// POUs/_FB_VisuDelta
(****************************************************************************************************<br>
© Syntegon Group.<br>
All rights reserved, also regarding any disposal, exploitation, reproduction, editing, distribution,<br>
as well as in the event of applications for industrial property rights.<br>
*****************************************************************************************************<br>
DESCRIPTION:<br>
One visualised Delta robot. Typical cycle:<br>
  fb_Delta.m_Register(vio_Manifest := GVL_Visu.stManifest, vi_udn_Id := 10, vi_str_Name := 'Delta 1',<br>
      vi_str_Path := 'MAIN.fb_Delta.vo_Visu');<br>
  fb_Delta.m_Configure(vi_Pose := BasePose, vi_lr_BaseRadius := 200, vi_lr_EffectorRadius := 50,<br>
      vi_lr_UpperArmLength := 400, vi_lr_LowerArmLength := 1000);<br>
  fb_Delta.m_SetFinger(vi_un_Finger := 1, vi_lr_Diameter := 40, vi_lr_Height := 50);<br>
  fb_Delta.m_SetWorkingArea(vi_lr_Radius := 750, vi_lr_ZMin := -1300, vi_lr_ZMax := -700, vi_lr_ConeHeight := 200,<br>
      vi_lr_ConeBottomRadius := 450);<br>
  fb_Delta.m_SetLimitArea(vi_lr_XMin := -500, vi_lr_XMax := 500, vi_lr_YMin := -750, vi_lr_YMax := 750,<br>
      vi_lr_ZMin := -1500, vi_lr_ZMax := -700);<br>
  fb_Delta.m_SetZone(vi_un_Zone := 1, vi_udn_ConveyorId := 1, vi_lr_Start := 1100, vi_lr_End := 1900,<br>
      vi_lr_AllocationOffset := 300);<br>
  fb_Delta.m_SetTcp(vi_ActualTcp := ActualTcp, vi_SetpointTcp := SetpointTcp);<br>
  fb_Delta.m_SetFingerState(vi_un_Finger := 1, vi_Pose := CupPose, vi_b_Active := b_Vacuum);<br>
Only the TCP (the gripper flange) is reported; the visualisation derives the arms from it. Tool rotations<br>
(e.g. a 4th axis) show only through the finger poses, absolute in the MCS. The config methods may be called<br>
every cycle; the config version only changes when a value does.<br>
*****************************************************************************************************<br>
OUTPUT VALUES:<br>
vo_Visu is the contract structure the gateway reads at the path given to m_Register. Do not write it.<br>
*****************************************************************************************************<br>
VERSION         ¦ DATE       ¦ NAME      ¦ CHANGE<br>
Syn_Visu 3.0.0  ¦ 2026-10-31 ¦ J.Willner ¦ Naming and layout after the TCAT programming guideline<br>
Syn_Visu 4.0.0  ¦ 2026-11-01 ¦ J.Willner ¦ Zones and fingers from _FB_VisuRobot; m_SetZone by index, no kind<br>
****************************************************************************************************)
FUNCTION_BLOCK _FB_VisuDelta EXTENDS _FB_VisuRobot
VAR_OUTPUT
	vo_Visu								: ST_VisuDelta;	// contract structure read by the gateway
END_VAR

(****************************************************************************************************<br>
© Syntegon Group.<br>
All rights reserved, also regarding any disposal, exploitation, reproduction, editing, distribution,<br>
as well as in the event of applications for industrial property rights.<br>
*****************************************************************************************************<br>
DESCRIPTION:<br>
Takes over vio_New and increments the config version if it differs from the current config. TRUE if changed.<br>
****************************************************************************************************)
METHOD PRIVATE m_ApplyConfig : BOOL
VAR_IN_OUT
	vio_New								: ST_VisuDeltaConfig;
END_VAR
m_ApplyConfig := Tc2_System.MEMCMP(ADR(vio_New), ADR(vo_Visu.stConfig), SIZEOF(vio_New)) <> 0;
IF m_ApplyConfig THEN
	vo_Visu.stConfig := vio_New;
	m_NotifyConfigChanged();
END_IF
END_METHOD

(****************************************************************************************************<br>
© Syntegon Group.<br>
All rights reserved, also regarding any disposal, exploitation, reproduction, editing, distribution,<br>
as well as in the event of applications for industrial property rights.<br>
*****************************************************************************************************<br>
DESCRIPTION:<br>
Base pose last set by m_Configure, MCS.<br>
****************************************************************************************************)
METHOD m_BasePose : ST_VisuPose
m_BasePose := vo_Visu.stConfig.stPose;
END_METHOD

(****************************************************************************************************<br>
© Syntegon Group.<br>
All rights reserved, also regarding any disposal, exploitation, reproduction, editing, distribution,<br>
as well as in the event of applications for industrial property rights.<br>
*****************************************************************************************************<br>
DESCRIPTION:<br>
Removes the limit area. TRUE if changed.<br>
****************************************************************************************************)
METHOD m_ClearLimitArea : BOOL
VAR
	TempNew								: ST_VisuDeltaConfig;
	TempEmpty							: ST_VisuLimitArea;
END_VAR
TempNew := vo_Visu.stConfig;
TempNew.stLimitArea := TempEmpty;
m_ClearLimitArea := m_ApplyConfig(TempNew);
END_METHOD

(****************************************************************************************************<br>
© Syntegon Group.<br>
All rights reserved, also regarding any disposal, exploitation, reproduction, editing, distribution,<br>
as well as in the event of applications for industrial property rights.<br>
*****************************************************************************************************<br>
DESCRIPTION:<br>
Manifest type: Delta robot.<br>
****************************************************************************************************)
METHOD PROTECTED m_ComponentType : E_VisuComponentType
m_ComponentType := E_VisuComponentType.DELTA;
END_METHOD

(****************************************************************************************************<br>
© Syntegon Group.<br>
All rights reserved, also regarding any disposal, exploitation, reproduction, editing, distribution,<br>
as well as in the event of applications for industrial property rights.<br>
*****************************************************************************************************<br>
DESCRIPTION:<br>
Sets base pose and geometry. Arm 1 lies along the base's local +X; arms 2 and 3 follow<br>
counter-clockwise (seen from above) at 120 deg each. TRUE if anything changed.<br>
****************************************************************************************************)
METHOD m_Configure : BOOL
VAR_INPUT
	vi_Pose								: ST_VisuPose;	// MCS, base centre
	vi_lr_BaseRadius					: LREAL;	// [mm] base centre to shoulder joint
	vi_lr_EffectorRadius				: LREAL;	// [mm] effector centre to lower-arm joint
	vi_lr_UpperArmLength				: LREAL;	// [mm]
	vi_lr_LowerArmLength				: LREAL;	// [mm]
END_VAR
VAR
	TempNew								: ST_VisuDeltaConfig;
END_VAR
TempNew := vo_Visu.stConfig;
TempNew.stPose := vi_Pose;
TempNew.fBaseRadius := vi_lr_BaseRadius;
TempNew.fEffectorRadius := vi_lr_EffectorRadius;
TempNew.fUpperArmLength := vi_lr_UpperArmLength;
TempNew.fLowerArmLength := vi_lr_LowerArmLength;
m_Configure := m_ApplyConfig(TempNew);
END_METHOD

(****************************************************************************************************<br>
© Syntegon Group.<br>
All rights reserved, also regarding any disposal, exploitation, reproduction, editing, distribution,<br>
as well as in the event of applications for industrial property rights.<br>
*****************************************************************************************************<br>
DESCRIPTION:<br>
The robot's gripper fingers for _FB_VisuRobot.m_SetFinger and m_ClearFingers.<br>
****************************************************************************************************)
METHOD PROTECTED m_Fingers : BOOL
VAR_OUTPUT
	vo_p_Count							: POINTER TO UINT;
	vo_p_Fingers						: POINTER TO ARRAY[0..VISU_GlobalConst_Param.VISU_un_MAX_FINGERS - 1] OF ST_VisuFinger;
END_VAR
vo_p_Count := ADR(vo_Visu.stConfig.nFingerCount);
vo_p_Fingers := ADR(vo_Visu.stConfig.aFingers);
m_Fingers := TRUE;
END_METHOD

(****************************************************************************************************<br>
© Syntegon Group.<br>
All rights reserved, also regarding any disposal, exploitation, reproduction, editing, distribution,<br>
as well as in the event of applications for industrial property rights.<br>
*****************************************************************************************************<br>
DESCRIPTION:<br>
Sets or clears the fault of the robot: drawn red with the message while active. The fault stays until it<br>
is cleared with m_SetFault(vi_b_Active := FALSE, vi_str_Message := ''). TRUE.<br>
****************************************************************************************************)
METHOD m_SetFault : BOOL
VAR_INPUT
	vi_b_Active							: BOOL;	// TRUE: fault active
	vi_str_Message						: STRING(80);	// shown to the operator; empty shows 'Fault'
END_VAR
vo_Visu.stState.stFault.bActive := vi_b_Active;
vo_Visu.stState.stFault.sMessage := vi_str_Message;
m_SetFault := TRUE;
END_METHOD

(****************************************************************************************************<br>
© Syntegon Group.<br>
All rights reserved, also regarding any disposal, exploitation, reproduction, editing, distribution,<br>
as well as in the event of applications for industrial property rights.<br>
*****************************************************************************************************<br>
DESCRIPTION:<br>
Reports finger vi_un_Finger (1-based): the pose of its frame (centre of its top face), absolute in the MCS,<br>
and whether it grips. Call once per cycle per configured finger.<br>
*****************************************************************************************************<br>
OUTPUT VALUES:<br>
FALSE outside 1..VISU_GlobalConst_Param.VISU_un_MAX_FINGERS.<br>
****************************************************************************************************)
METHOD m_SetFingerState : BOOL
VAR_INPUT
	vi_un_Finger						: UINT;	// [-] 1-based
	vi_Pose								: ST_VisuPose;	// MCS
	vi_b_Active							: BOOL;	// TRUE while the finger grips
END_VAR
m_SetFingerState := vi_un_Finger > 0 AND vi_un_Finger <= VISU_GlobalConst_Param.VISU_un_MAX_FINGERS;
IF m_SetFingerState THEN
	vo_Visu.stState.aFingerStates[vi_un_Finger - 1].stPose := vi_Pose;
	vo_Visu.stState.aFingerStates[vi_un_Finger - 1].bActive := vi_b_Active;
END_IF
END_METHOD

(****************************************************************************************************<br>
© Syntegon Group.<br>
All rights reserved, also regarding any disposal, exploitation, reproduction, editing, distribution,<br>
as well as in the event of applications for industrial property rights.<br>
*****************************************************************************************************<br>
DESCRIPTION:<br>
Sets and activates the limit area: an axis-aligned box in the robot frame. TRUE if changed.<br>
****************************************************************************************************)
METHOD m_SetLimitArea : BOOL
VAR_INPUT
	vi_lr_XMin							: LREAL;	// [mm]
	vi_lr_XMax							: LREAL;	// [mm]
	vi_lr_YMin							: LREAL;	// [mm]
	vi_lr_YMax							: LREAL;	// [mm]
	vi_lr_ZMin							: LREAL;	// [mm] relative to the base (below the base: negative)
	vi_lr_ZMax							: LREAL;	// [mm] relative to the base
END_VAR
VAR
	TempNew								: ST_VisuDeltaConfig;
END_VAR
TempNew := vo_Visu.stConfig;
TempNew.stLimitArea.fXMin := vi_lr_XMin;
TempNew.stLimitArea.fXMax := vi_lr_XMax;
TempNew.stLimitArea.fYMin := vi_lr_YMin;
TempNew.stLimitArea.fYMax := vi_lr_YMax;
TempNew.stLimitArea.fZMin := vi_lr_ZMin;
TempNew.stLimitArea.fZMax := vi_lr_ZMax;
TempNew.stLimitArea.bActive := TRUE;
m_SetLimitArea := m_ApplyConfig(TempNew);
END_METHOD

(****************************************************************************************************<br>
© Syntegon Group.<br>
All rights reserved, also regarding any disposal, exploitation, reproduction, editing, distribution,<br>
as well as in the event of applications for industrial property rights.<br>
*****************************************************************************************************<br>
DESCRIPTION:<br>
Moves the robot's shown coordinate system (origin triad, local measuring coordinates) away from the base<br>
centre (stPose), in the base's local frame. Geometry, working area and limit area stay relative to stPose.<br>
TRUE if anything changed.<br>
****************************************************************************************************)
METHOD m_SetOriginShift : BOOL
VAR_INPUT
	vi_lr_X								: LREAL;	// [mm] along the base's local X
	vi_lr_Y								: LREAL := 0;	// [mm] along the base's local Y
	vi_lr_Z								: LREAL := 0;	// [mm] along the base's local Z
END_VAR
VAR
	TempNew								: ST_VisuDeltaConfig;
END_VAR
TempNew := vo_Visu.stConfig;
TempNew.stOriginShift.fX := vi_lr_X;
TempNew.stOriginShift.fY := vi_lr_Y;
TempNew.stOriginShift.fZ := vi_lr_Z;
m_SetOriginShift := m_ApplyConfig(TempNew);
END_METHOD

(****************************************************************************************************<br>
© Syntegon Group.<br>
All rights reserved, also regarding any disposal, exploitation, reproduction, editing, distribution,<br>
as well as in the event of applications for industrial property rights.<br>
*****************************************************************************************************<br>
DESCRIPTION:<br>
Reports the robot's TCP. Call once per cycle; it also stamps the state with the cycle's DC time.<br>
****************************************************************************************************)
METHOD m_SetTcp : BOOL
VAR_INPUT
	vi_ActualTcp						: ST_VisuPosition;	// MCS, effector centre (the gripper flange)
	vi_SetpointTcp						: ST_VisuPosition;	// MCS
END_VAR
vo_Visu.stState.stActualTcp := vi_ActualTcp;
vo_Visu.stState.stSetpointTcp := vi_SetpointTcp;
vo_Visu.stState.nTimestamp := m_DcTime();
m_SetTcp := TRUE;
END_METHOD

(****************************************************************************************************<br>
© Syntegon Group.<br>
All rights reserved, also regarding any disposal, exploitation, reproduction, editing, distribution,<br>
as well as in the event of applications for industrial property rights.<br>
*****************************************************************************************************<br>
DESCRIPTION:<br>
Sets the working area: a vertical cylinder in the robot frame with an optional cone below. TRUE if changed.<br>
****************************************************************************************************)
METHOD m_SetWorkingArea : BOOL
VAR_INPUT
	vi_lr_Radius						: LREAL;	// [mm]
	vi_lr_ZMin							: LREAL;	// [mm] relative to the base (below the base: negative)
	vi_lr_ZMax							: LREAL;	// [mm] relative to the base
	vi_lr_ConeHeight					: LREAL;	// [mm] below vi_lr_ZMin; 0 = no cone
	vi_lr_ConeBottomRadius				: LREAL;	// [mm]
END_VAR
VAR
	TempNew								: ST_VisuDeltaConfig;
END_VAR
TempNew := vo_Visu.stConfig;
TempNew.stWorkingArea.fRadius := vi_lr_Radius;
TempNew.stWorkingArea.fZMin := vi_lr_ZMin;
TempNew.stWorkingArea.fZMax := vi_lr_ZMax;
TempNew.stWorkingArea.fConeHeight := vi_lr_ConeHeight;
TempNew.stWorkingArea.fConeBottomRadius := vi_lr_ConeBottomRadius;
m_SetWorkingArea := m_ApplyConfig(TempNew);
END_METHOD

(****************************************************************************************************<br>
© Syntegon Group.<br>
All rights reserved, also regarding any disposal, exploitation, reproduction, editing, distribution,<br>
as well as in the event of applications for industrial property rights.<br>
*****************************************************************************************************<br>
DESCRIPTION:<br>
The robot's zones for _FB_VisuZoneComponent.m_SetZone and m_ClearZones.<br>
****************************************************************************************************)
METHOD PROTECTED m_Zones : BOOL
VAR_OUTPUT
	vo_p_Count							: POINTER TO UINT;
	vo_p_Zones							: POINTER TO ARRAY[0..VISU_GlobalConst_Param.VISU_un_MAX_ZONES - 1] OF ST_VisuZone;
END_VAR
vo_p_Count := ADR(vo_Visu.stConfig.nZoneCount);
vo_p_Zones := ADR(vo_Visu.stConfig.aZones);
m_Zones := TRUE;
END_METHOD

END_FUNCTION_BLOCK

// POUs/_FB_VisuRobot
(****************************************************************************************************<br>
© Syntegon Group.<br>
All rights reserved, also regarding any disposal, exploitation, reproduction, editing, distribution,<br>
as well as in the event of applications for industrial property rights.<br>
*****************************************************************************************************<br>
DESCRIPTION:<br>
Base of every robot (Delta, XTS gantry, XTS loop, Cartesian): zones plus the gripper fingers,<br>
m_SetFinger and m_ClearFingers. A derived FB tells where its fingers lie through m_Fingers.<br>
Not used directly.<br>
*****************************************************************************************************<br>
VERSION         ¦ DATE       ¦ NAME      ¦ CHANGE<br>
Syn_Visu 4.0.0  ¦ 2026-11-01 ¦ J.Willner ¦ New: fingers shared by all robots<br>
****************************************************************************************************)
FUNCTION_BLOCK ABSTRACT _FB_VisuRobot EXTENDS _FB_VisuZoneComponent

(****************************************************************************************************<br>
© Syntegon Group.<br>
All rights reserved, also regarding any disposal, exploitation, reproduction, editing, distribution,<br>
as well as in the event of applications for industrial property rights.<br>
*****************************************************************************************************<br>
DESCRIPTION:<br>
Removes the gripper definition. TRUE if there was one.<br>
****************************************************************************************************)
METHOD m_ClearFingers : BOOL
VAR
	p_TempCount							: POINTER TO UINT;
	p_TempFingers						: POINTER TO ARRAY[0..VISU_GlobalConst_Param.VISU_un_MAX_FINGERS - 1] OF ST_VisuFinger;
	TempEmpty							: ST_VisuFinger;
	un_TempIndex						: UINT;
END_VAR
m_ClearFingers := FALSE;
m_Fingers(vo_p_Count => p_TempCount, vo_p_Fingers => p_TempFingers);
IF p_TempCount = 0 OR p_TempFingers = 0 THEN
	RETURN;
END_IF
m_ClearFingers := p_TempCount^ > 0;
FOR un_TempIndex := 0 TO VISU_GlobalConst_Param.VISU_un_MAX_FINGERS - 1 DO
	p_TempFingers^[un_TempIndex] := TempEmpty;
END_FOR
p_TempCount^ := 0;
IF m_ClearFingers THEN
	m_NotifyConfigChanged();
END_IF
END_METHOD

(****************************************************************************************************<br>
© Syntegon Group.<br>
All rights reserved, also regarding any disposal, exploitation, reproduction, editing, distribution,<br>
as well as in the event of applications for industrial property rights.<br>
*****************************************************************************************************<br>
DESCRIPTION:<br>
Where the gripper fingers lie in the derived FB's contract structure: vo_p_Count points to its<br>
nFingerCount, vo_p_Fingers to its aFingers.<br>
****************************************************************************************************)
METHOD PROTECTED ABSTRACT m_Fingers : BOOL
VAR_OUTPUT
	vo_p_Count							: POINTER TO UINT;
	vo_p_Fingers						: POINTER TO ARRAY[0..VISU_GlobalConst_Param.VISU_un_MAX_FINGERS - 1] OF ST_VisuFinger;
END_VAR
END_METHOD

(****************************************************************************************************<br>
© Syntegon Group.<br>
All rights reserved, also regarding any disposal, exploitation, reproduction, editing, distribution,<br>
as well as in the event of applications for industrial property rights.<br>
*****************************************************************************************************<br>
DESCRIPTION:<br>
Defines gripper finger vi_un_Finger (1-based): a cylinder hanging from the finger's pose along its local -Z.<br>
For XTS kinematics it is a finger of every mover's gripper. The finger count grows to vi_un_Finger.<br>
*****************************************************************************************************<br>
OUTPUT VALUES:<br>
FALSE outside 1..VISU_GlobalConst_Param.VISU_un_MAX_FINGERS.<br>
****************************************************************************************************)
METHOD m_SetFinger : BOOL
VAR_INPUT
	vi_un_Finger						: UINT;	// [-] 1-based, as a product's nFingerId
	vi_lr_Diameter						: LREAL;	// [mm]
	vi_lr_Height						: LREAL;	// [mm] along the finger's local -Z
END_VAR
VAR
	p_TempCount							: POINTER TO UINT;
	p_TempFingers						: POINTER TO ARRAY[0..VISU_GlobalConst_Param.VISU_un_MAX_FINGERS - 1] OF ST_VisuFinger;
	TempFinger							: ST_VisuFinger;
END_VAR
m_SetFinger := FALSE;
IF vi_un_Finger = 0 OR vi_un_Finger > VISU_GlobalConst_Param.VISU_un_MAX_FINGERS THEN
	RETURN;
END_IF
m_Fingers(vo_p_Count => p_TempCount, vo_p_Fingers => p_TempFingers);
IF p_TempCount = 0 OR p_TempFingers = 0 THEN
	RETURN;
END_IF
TempFinger.fDiameter := vi_lr_Diameter;
TempFinger.fHeight := vi_lr_Height;
IF vi_un_Finger > p_TempCount^
OR Tc2_System.MEMCMP(ADR(TempFinger), ADR(p_TempFingers^[vi_un_Finger - 1]), SIZEOF(TempFinger)) <> 0
THEN
	p_TempFingers^[vi_un_Finger - 1] := TempFinger;
	p_TempCount^ := MAX(p_TempCount^, vi_un_Finger);
	m_NotifyConfigChanged();
END_IF
m_SetFinger := TRUE;
END_METHOD

END_FUNCTION_BLOCK

// POUs/_FB_VisuZoneComponent
(****************************************************************************************************<br>
© Syntegon Group.<br>
All rights reserved, also regarding any disposal, exploitation, reproduction, editing, distribution,<br>
as well as in the event of applications for industrial property rights.<br>
*****************************************************************************************************<br>
DESCRIPTION:<br>
Base of every component with zones on conveyors (robots, detectors): m_SetZone and m_ClearZones.<br>
A derived FB tells where its zones lie in its contract structure through m_Zones. Not used directly.<br>
*****************************************************************************************************<br>
VERSION         ¦ DATE       ¦ NAME      ¦ CHANGE<br>
Syn_Visu 4.0.0  ¦ 2026-11-01 ¦ J.Willner ¦ New: zones shared by robots and detectors, no zone kind<br>
****************************************************************************************************)
FUNCTION_BLOCK ABSTRACT _FB_VisuZoneComponent EXTENDS _FB_VisuComponent

(****************************************************************************************************<br>
© Syntegon Group.<br>
All rights reserved, also regarding any disposal, exploitation, reproduction, editing, distribution,<br>
as well as in the event of applications for industrial property rights.<br>
*****************************************************************************************************<br>
DESCRIPTION:<br>
Removes all zones. TRUE if there were any.<br>
****************************************************************************************************)
METHOD m_ClearZones : BOOL
VAR
	p_TempCount							: POINTER TO UINT;
	p_TempZones							: POINTER TO ARRAY[0..VISU_GlobalConst_Param.VISU_un_MAX_ZONES - 1] OF ST_VisuZone;
	TempEmpty							: ST_VisuZone;
	un_TempIndex						: UINT;
END_VAR
m_ClearZones := FALSE;
m_Zones(vo_p_Count => p_TempCount, vo_p_Zones => p_TempZones);
IF p_TempCount = 0 OR p_TempZones = 0 THEN
	RETURN;
END_IF
m_ClearZones := p_TempCount^ > 0;
FOR un_TempIndex := 0 TO VISU_GlobalConst_Param.VISU_un_MAX_ZONES - 1 DO
	p_TempZones^[un_TempIndex] := TempEmpty;
END_FOR
p_TempCount^ := 0;
IF m_ClearZones THEN
	m_NotifyConfigChanged();
END_IF
END_METHOD

(****************************************************************************************************<br>
© Syntegon Group.<br>
All rights reserved, also regarding any disposal, exploitation, reproduction, editing, distribution,<br>
as well as in the event of applications for industrial property rights.<br>
*****************************************************************************************************<br>
DESCRIPTION:<br>
Sets zone vi_un_Zone (1-based): a stretch of a conveyor that belongs to this component, e.g. where a<br>
robot picks or places or where a detector detects. vi_lr_Start = vi_lr_End is a line across the belt.<br>
The zone count grows to vi_un_Zone; set the zones in order. The config version only changes when a<br>
value does.<br>
*****************************************************************************************************<br>
OUTPUT VALUES:<br>
FALSE for vi_udn_ConveyorId = 0 or vi_un_Zone outside 1..VISU_GlobalConst_Param.VISU_un_MAX_ZONES.<br>
****************************************************************************************************)
METHOD m_SetZone : BOOL
VAR_INPUT
	vi_un_Zone							: UINT;	// [-] 1-based
	vi_udn_ConveyorId					: UDINT;	// [-] manifest id of the conveyor
	vi_lr_Start							: LREAL;	// [mm] along the conveyor from its origin (belt coordinates, not MCS)
	vi_lr_End							: LREAL;	// [mm] along the conveyor from its origin
	vi_lr_AllocationOffset				: LREAL := 0;	// [mm] before vi_lr_End up to which products may be allocated; 0 = no limit
	vi_lr_CcsOffset						: LREAL := 0;	// [mm] along the conveyor from its origin: the component's conveyor coordinate system
END_VAR
VAR
	p_TempCount							: POINTER TO UINT;
	p_TempZones							: POINTER TO ARRAY[0..VISU_GlobalConst_Param.VISU_un_MAX_ZONES - 1] OF ST_VisuZone;
	TempZone							: ST_VisuZone;
END_VAR
m_SetZone := FALSE;
IF vi_udn_ConveyorId = 0 OR vi_un_Zone = 0 OR vi_un_Zone > VISU_GlobalConst_Param.VISU_un_MAX_ZONES THEN
	RETURN;
END_IF
m_Zones(vo_p_Count => p_TempCount, vo_p_Zones => p_TempZones);
IF p_TempCount = 0 OR p_TempZones = 0 THEN
	RETURN;
END_IF
TempZone.nConveyorId := vi_udn_ConveyorId;
TempZone.fStart := vi_lr_Start;
TempZone.fEnd := vi_lr_End;
TempZone.fAllocationOffset := vi_lr_AllocationOffset;
TempZone.fCcsOffset := vi_lr_CcsOffset;
IF vi_un_Zone > p_TempCount^
OR Tc2_System.MEMCMP(ADR(TempZone), ADR(p_TempZones^[vi_un_Zone - 1]), SIZEOF(TempZone)) <> 0
THEN
	p_TempZones^[vi_un_Zone - 1] := TempZone;
	p_TempCount^ := MAX(p_TempCount^, vi_un_Zone);
	m_NotifyConfigChanged();
END_IF
m_SetZone := TRUE;
END_METHOD

(****************************************************************************************************<br>
© Syntegon Group.<br>
All rights reserved, also regarding any disposal, exploitation, reproduction, editing, distribution,<br>
as well as in the event of applications for industrial property rights.<br>
*****************************************************************************************************<br>
DESCRIPTION:<br>
Where the zones lie in the derived FB's contract structure: vo_p_Count points to its nZoneCount,<br>
vo_p_Zones to its aZones.<br>
****************************************************************************************************)
METHOD PROTECTED ABSTRACT m_Zones : BOOL
VAR_OUTPUT
	vo_p_Count							: POINTER TO UINT;
	vo_p_Zones							: POINTER TO ARRAY[0..VISU_GlobalConst_Param.VISU_un_MAX_ZONES - 1] OF ST_VisuZone;
END_VAR
END_METHOD

END_FUNCTION_BLOCK

// POUs/_FB_VisuStation
(****************************************************************************************************<br>
© Syntegon Group.<br>
All rights reserved, also regarding any disposal, exploitation, reproduction, editing, distribution,<br>
as well as in the event of applications for industrial property rights.<br>
*****************************************************************************************************<br>
DESCRIPTION:<br>
One visualised station: a client at a conveyor that works on the products in its zones, e.g. a reject<br>
unit, a labeller, a printer or a check weigher. It is drawn only from the bodies it describes. Typical cycle<br>
of a reject unit:<br>
  fb_Reject.m_Register(vio_Manifest := GVL_Visu.stManifest, vi_udn_Id := 70, vi_str_Name := 'Reject unit',<br>
      vi_str_Path := 'MAIN.fb_Reject.vo_Visu');<br>
  fb_Reject.m_Configure(vi_Pose := StationPose);<br>
  fb_Reject.m_SetBody(vi_un_Body := 1, ...);   // housing<br>
  fb_Reject.m_SetBody(vi_un_Body := 2, ...);   // pusher<br>
  fb_Reject.m_SetZone(vi_un_Zone := 1, vi_udn_ConveyorId := 2, vi_lr_Start := 2400, vi_lr_End := 2400);<br>
  fb_Reject.m_SetBodyActive(vi_un_Body := 2, vi_b_Active := b_Pushing);<br>
and on the conveyor, when it rejects a product:<br>
  fb_Outfeed.m_SetProductState(vi_udn_Id := udn_Product, vi_e_State := E_VisuProductState.REJECTED,<br>
      vi_udn_ClientId := fb_Reject.m_Id());<br>
A station may also latch products (m_LatchProduct with vi_udn_ClientId := its id), e.g. a check weigher.<br>
*****************************************************************************************************<br>
OUTPUT VALUES:<br>
vo_Visu is the contract structure the gateway reads at the path given to m_Register. Do not write it.<br>
*****************************************************************************************************<br>
VERSION         ¦ DATE       ¦ NAME      ¦ CHANGE<br>
Syn_Visu 6.0.0  ¦ 2026-11-01 ¦ J.Willner ¦ New<br>
****************************************************************************************************)
FUNCTION_BLOCK _FB_VisuStation EXTENDS _FB_VisuBodyComponent
VAR_OUTPUT
	vo_Visu								: ST_VisuStation;	// contract structure read by the gateway
END_VAR

(****************************************************************************************************<br>
© Syntegon Group.<br>
All rights reserved, also regarding any disposal, exploitation, reproduction, editing, distribution,<br>
as well as in the event of applications for industrial property rights.<br>
*****************************************************************************************************<br>
DESCRIPTION:<br>
Manifest type: station.<br>
****************************************************************************************************)
METHOD PROTECTED m_ComponentType : E_VisuComponentType
m_ComponentType := E_VisuComponentType.STATION;
END_METHOD

(****************************************************************************************************<br>
© Syntegon Group.<br>
All rights reserved, also regarding any disposal, exploitation, reproduction, editing, distribution,<br>
as well as in the event of applications for industrial property rights.<br>
*****************************************************************************************************<br>
DESCRIPTION:<br>
Sets the station's pose; its bodies (m_SetBody) are placed relative to it. TRUE if it changed.<br>
****************************************************************************************************)
METHOD m_Configure : BOOL
VAR_INPUT
	vi_Pose								: ST_VisuPose;	// MCS, the station's origin, e.g. at the belt side on the floor
END_VAR
m_Configure := m_SetPose(vi_Pose);
END_METHOD

(****************************************************************************************************<br>
© Syntegon Group.<br>
All rights reserved, also regarding any disposal, exploitation, reproduction, editing, distribution,<br>
as well as in the event of applications for industrial property rights.<br>
*****************************************************************************************************<br>
DESCRIPTION:<br>
The station's pose, origin shift, bodies, body states, timestamp and fault for _FB_VisuBodyComponent.<br>
****************************************************************************************************)
METHOD PROTECTED m_Parts : BOOL
VAR_OUTPUT
	vo_p_Pose							: POINTER TO ST_VisuPose;
	vo_p_OriginShift					: POINTER TO ST_VisuPosition;
	vo_p_BodyCount						: POINTER TO UINT;
	vo_p_Bodies							: POINTER TO ARRAY[0..VISU_GlobalConst_Param.VISU_un_MAX_BODIES - 1] OF ST_VisuBody;
	vo_p_BodyStates						: POINTER TO ARRAY[0..VISU_GlobalConst_Param.VISU_un_MAX_BODIES - 1] OF ST_VisuBodyState;
	vo_p_Timestamp						: POINTER TO ULINT;
	vo_p_Fault							: POINTER TO ST_VisuFault;
END_VAR
vo_p_Pose := ADR(vo_Visu.stConfig.stPose);
vo_p_OriginShift := ADR(vo_Visu.stConfig.stOriginShift);
vo_p_BodyCount := ADR(vo_Visu.stConfig.nBodyCount);
vo_p_Bodies := ADR(vo_Visu.stConfig.aBodies);
vo_p_BodyStates := ADR(vo_Visu.stState.aBodyStates);
vo_p_Timestamp := ADR(vo_Visu.stState.nTimestamp);
vo_p_Fault := ADR(vo_Visu.stState.stFault);
m_Parts := TRUE;
END_METHOD

(****************************************************************************************************<br>
© Syntegon Group.<br>
All rights reserved, also regarding any disposal, exploitation, reproduction, editing, distribution,<br>
as well as in the event of applications for industrial property rights.<br>
*****************************************************************************************************<br>
DESCRIPTION:<br>
The station's zones for _FB_VisuZoneComponent.m_SetZone and m_ClearZones.<br>
****************************************************************************************************)
METHOD PROTECTED m_Zones : BOOL
VAR_OUTPUT
	vo_p_Count							: POINTER TO UINT;
	vo_p_Zones							: POINTER TO ARRAY[0..VISU_GlobalConst_Param.VISU_un_MAX_ZONES - 1] OF ST_VisuZone;
END_VAR
vo_p_Count := ADR(vo_Visu.stConfig.nZoneCount);
vo_p_Zones := ADR(vo_Visu.stConfig.aZones);
m_Zones := TRUE;
END_METHOD

END_FUNCTION_BLOCK

// POUs/_FB_VisuCartesian
(****************************************************************************************************<br>
© Syntegon Group.<br>
All rights reserved, also regarding any disposal, exploitation, reproduction, editing, distribution,<br>
as well as in the event of applications for industrial property rights.<br>
*****************************************************************************************************<br>
DESCRIPTION:<br>
One visualised Cartesian robot: linear X, Y, Z axes ending at a gripper flange. Typical cycle:<br>
  fb_Cartesian.m_Register(vio_Manifest := GVL_Visu.stManifest, vi_udn_Id := 40, vi_str_Name := 'Cartesian',<br>
      vi_str_Path := 'MAIN.fb_Cartesian.vo_Visu');<br>
  fb_Cartesian.m_Configure(vi_Pose := RobotPose, vi_lr_XMin := 0, vi_lr_XMax := 1200, vi_lr_YMin := 0,<br>
      vi_lr_YMax := 1000, vi_lr_ZMin := -600, vi_lr_ZMax := 0, vi_lr_RailHeight := 1200);<br>
  fb_Cartesian.m_SetFinger(vi_un_Finger := 1, vi_lr_Diameter := 40, vi_lr_Height := 40);<br>
  fb_Cartesian.m_SetZone(vi_un_Zone := 1, vi_udn_ConveyorId := 7, vi_lr_Start := 1000, vi_lr_End := 2000);<br>
  fb_Cartesian.m_SetAxes(vi_lr_X := ..., vi_lr_Y := ..., vi_lr_Z := ...);<br>
  fb_Cartesian.m_SetFingerState(vi_un_Finger := 1, vi_Pose := CupPose, vi_b_Active := b_Vacuum);<br>
Only actual values are reported; tool rotations (e.g. C and A) show only through the finger poses, absolute in<br>
the MCS. The config methods may be called every cycle; the config version only changes when a value does.<br>
*****************************************************************************************************<br>
OUTPUT VALUES:<br>
vo_Visu is the contract structure the gateway reads at the path given to m_Register. Do not write it.<br>
*****************************************************************************************************<br>
VERSION         ¦ DATE       ¦ NAME      ¦ CHANGE<br>
Syn_Visu 3.0.0  ¦ 2026-10-31 ¦ J.Willner ¦ Naming and layout after the TCAT programming guideline<br>
Syn_Visu 4.0.0  ¦ 2026-11-01 ¦ J.Willner ¦ Zones and fingers from _FB_VisuRobot; m_SetZone by index, no kind<br>
****************************************************************************************************)
FUNCTION_BLOCK _FB_VisuCartesian EXTENDS _FB_VisuRobot
VAR_OUTPUT
	vo_Visu								: ST_VisuCartesian;	// contract structure read by the gateway
END_VAR

(****************************************************************************************************<br>
© Syntegon Group.<br>
All rights reserved, also regarding any disposal, exploitation, reproduction, editing, distribution,<br>
as well as in the event of applications for industrial property rights.<br>
*****************************************************************************************************<br>
DESCRIPTION:<br>
Takes over vio_New and increments the config version if it differs from the current config. TRUE if changed.<br>
****************************************************************************************************)
METHOD PRIVATE m_ApplyConfig : BOOL
VAR_IN_OUT
	vio_New								: ST_VisuCartesianConfig;
END_VAR
m_ApplyConfig := Tc2_System.MEMCMP(ADR(vio_New), ADR(vo_Visu.stConfig), SIZEOF(vio_New)) <> 0;
IF m_ApplyConfig THEN
	vo_Visu.stConfig := vio_New;
	m_NotifyConfigChanged();
END_IF
END_METHOD

(****************************************************************************************************<br>
© Syntegon Group.<br>
All rights reserved, also regarding any disposal, exploitation, reproduction, editing, distribution,<br>
as well as in the event of applications for industrial property rights.<br>
*****************************************************************************************************<br>
DESCRIPTION:<br>
Manifest type: Cartesian robot.<br>
****************************************************************************************************)
METHOD PROTECTED m_ComponentType : E_VisuComponentType
m_ComponentType := E_VisuComponentType.CARTESIAN;
END_METHOD

(****************************************************************************************************<br>
© Syntegon Group.<br>
All rights reserved, also regarding any disposal, exploitation, reproduction, editing, distribution,<br>
as well as in the event of applications for industrial property rights.<br>
*****************************************************************************************************<br>
DESCRIPTION:<br>
Sets pose, strokes and rail height. TRUE if anything changed.<br>
****************************************************************************************************)
METHOD m_Configure : BOOL
VAR_INPUT
	vi_Pose								: ST_VisuPose;	// MCS, axis origin X = Y = 0 with Z up
	vi_lr_XMin							: LREAL;	// [mm]
	vi_lr_XMax							: LREAL;	// [mm]
	vi_lr_YMin							: LREAL;	// [mm]
	vi_lr_YMax							: LREAL;	// [mm]
	vi_lr_ZMin							: LREAL;	// [mm]
	vi_lr_ZMax							: LREAL;	// [mm]
	vi_lr_RailHeight					: LREAL;	// [mm] top of the rails above the local origin
END_VAR
VAR
	TempNew								: ST_VisuCartesianConfig;
END_VAR
TempNew := vo_Visu.stConfig;
TempNew.stPose := vi_Pose;
TempNew.fXMin := vi_lr_XMin;
TempNew.fXMax := vi_lr_XMax;
TempNew.fYMin := vi_lr_YMin;
TempNew.fYMax := vi_lr_YMax;
TempNew.fZMin := vi_lr_ZMin;
TempNew.fZMax := vi_lr_ZMax;
TempNew.fRailHeight := vi_lr_RailHeight;
m_Configure := m_ApplyConfig(TempNew);
END_METHOD

(****************************************************************************************************<br>
© Syntegon Group.<br>
All rights reserved, also regarding any disposal, exploitation, reproduction, editing, distribution,<br>
as well as in the event of applications for industrial property rights.<br>
*****************************************************************************************************<br>
DESCRIPTION:<br>
The robot's gripper fingers for _FB_VisuRobot.m_SetFinger and m_ClearFingers.<br>
****************************************************************************************************)
METHOD PROTECTED m_Fingers : BOOL
VAR_OUTPUT
	vo_p_Count							: POINTER TO UINT;
	vo_p_Fingers						: POINTER TO ARRAY[0..VISU_GlobalConst_Param.VISU_un_MAX_FINGERS - 1] OF ST_VisuFinger;
END_VAR
vo_p_Count := ADR(vo_Visu.stConfig.nFingerCount);
vo_p_Fingers := ADR(vo_Visu.stConfig.aFingers);
m_Fingers := TRUE;
END_METHOD

(****************************************************************************************************<br>
© Syntegon Group.<br>
All rights reserved, also regarding any disposal, exploitation, reproduction, editing, distribution,<br>
as well as in the event of applications for industrial property rights.<br>
*****************************************************************************************************<br>
DESCRIPTION:<br>
Reports the axes' actual values and the gripper. Call once per cycle; it also stamps the state with the<br>
cycle's DC time.<br>
****************************************************************************************************)
METHOD m_SetAxes : BOOL
VAR_INPUT
	vi_lr_X								: LREAL;	// [mm]
	vi_lr_Y								: LREAL;	// [mm]
	vi_lr_Z								: LREAL;	// [mm]
	vi_b_GripperActive					: BOOL := FALSE;	// used only when no fingers are configured
END_VAR
vo_Visu.stState.fX := vi_lr_X;
vo_Visu.stState.fY := vi_lr_Y;
vo_Visu.stState.fZ := vi_lr_Z;
vo_Visu.stState.bGripperActive := vi_b_GripperActive;
vo_Visu.stState.nTimestamp := m_DcTime();
m_SetAxes := TRUE;
END_METHOD

(****************************************************************************************************<br>
© Syntegon Group.<br>
All rights reserved, also regarding any disposal, exploitation, reproduction, editing, distribution,<br>
as well as in the event of applications for industrial property rights.<br>
*****************************************************************************************************<br>
DESCRIPTION:<br>
Sets or clears the fault of the robot: drawn red with the message while active. The fault stays until it<br>
is cleared with m_SetFault(vi_b_Active := FALSE, vi_str_Message := ''). TRUE.<br>
****************************************************************************************************)
METHOD m_SetFault : BOOL
VAR_INPUT
	vi_b_Active							: BOOL;	// TRUE: fault active
	vi_str_Message						: STRING(80);	// shown to the operator; empty shows 'Fault'
END_VAR
vo_Visu.stState.stFault.bActive := vi_b_Active;
vo_Visu.stState.stFault.sMessage := vi_str_Message;
m_SetFault := TRUE;
END_METHOD

(****************************************************************************************************<br>
© Syntegon Group.<br>
All rights reserved, also regarding any disposal, exploitation, reproduction, editing, distribution,<br>
as well as in the event of applications for industrial property rights.<br>
*****************************************************************************************************<br>
DESCRIPTION:<br>
Reports finger vi_un_Finger (1-based): the pose of its frame (centre of its top face), absolute in the MCS,<br>
and whether it grips. Call once per cycle per configured finger.<br>
*****************************************************************************************************<br>
OUTPUT VALUES:<br>
FALSE outside 1..VISU_GlobalConst_Param.VISU_un_MAX_FINGERS.<br>
****************************************************************************************************)
METHOD m_SetFingerState : BOOL
VAR_INPUT
	vi_un_Finger						: UINT;	// [-] 1-based
	vi_Pose								: ST_VisuPose;	// MCS
	vi_b_Active							: BOOL;	// TRUE while the finger grips
END_VAR
m_SetFingerState := vi_un_Finger > 0 AND vi_un_Finger <= VISU_GlobalConst_Param.VISU_un_MAX_FINGERS;
IF m_SetFingerState THEN
	vo_Visu.stState.aFingerStates[vi_un_Finger - 1].stPose := vi_Pose;
	vo_Visu.stState.aFingerStates[vi_un_Finger - 1].bActive := vi_b_Active;
END_IF
END_METHOD

(****************************************************************************************************<br>
© Syntegon Group.<br>
All rights reserved, also regarding any disposal, exploitation, reproduction, editing, distribution,<br>
as well as in the event of applications for industrial property rights.<br>
*****************************************************************************************************<br>
DESCRIPTION:<br>
Moves the robot's shown coordinate system (origin triad, local measuring coordinates) away from axis zero<br>
(stPose), in the robot's local frame. Geometry and axis values stay relative to stPose. TRUE if anything changed.<br>
****************************************************************************************************)
METHOD m_SetOriginShift : BOOL
VAR_INPUT
	vi_lr_X								: LREAL;	// [mm] along the robot's local X
	vi_lr_Y								: LREAL := 0;	// [mm] along the robot's local Y
	vi_lr_Z								: LREAL := 0;	// [mm] along the robot's local Z
END_VAR
VAR
	TempNew								: ST_VisuCartesianConfig;
END_VAR
TempNew := vo_Visu.stConfig;
TempNew.stOriginShift.fX := vi_lr_X;
TempNew.stOriginShift.fY := vi_lr_Y;
TempNew.stOriginShift.fZ := vi_lr_Z;
m_SetOriginShift := m_ApplyConfig(TempNew);
END_METHOD

(****************************************************************************************************<br>
© Syntegon Group.<br>
All rights reserved, also regarding any disposal, exploitation, reproduction, editing, distribution,<br>
as well as in the event of applications for industrial property rights.<br>
*****************************************************************************************************<br>
DESCRIPTION:<br>
The robot's zones for _FB_VisuZoneComponent.m_SetZone and m_ClearZones.<br>
****************************************************************************************************)
METHOD PROTECTED m_Zones : BOOL
VAR_OUTPUT
	vo_p_Count							: POINTER TO UINT;
	vo_p_Zones							: POINTER TO ARRAY[0..VISU_GlobalConst_Param.VISU_un_MAX_ZONES - 1] OF ST_VisuZone;
END_VAR
vo_p_Count := ADR(vo_Visu.stConfig.nZoneCount);
vo_p_Zones := ADR(vo_Visu.stConfig.aZones);
m_Zones := TRUE;
END_METHOD

END_FUNCTION_BLOCK

// POUs/_FB_VisuXtsGantry
(****************************************************************************************************<br>
© Syntegon Group.<br>
All rights reserved, also regarding any disposal, exploitation, reproduction, editing, distribution,<br>
as well as in the event of applications for industrial property rights.<br>
*****************************************************************************************************<br>
DESCRIPTION:<br>
One visualised XTS gantry (e.g. IDH): a straight track of XTS motor modules on a common Z axis, each mover<br>
with an X axis and a gripper flange at its end. Typical cycle:<br>
  fb_Idh.m_Register(vio_Manifest := GVL_Visu.stManifest, vi_udn_Id := 30, vi_str_Name := 'IDH',<br>
      vi_str_Path := 'MAIN.fb_Idh.vo_Visu');<br>
  fb_Idh.m_Configure(vi_Pose := TrackPose, vi_lr_XMin := 0, vi_lr_XMax := 700, vi_lr_ZMin := -100, vi_lr_ZMax := 0, vi_lr_ToolOffsetX := 150, vi_lr_ToolOffsetZ := -350,<br>
      vi_lr_MoverLength := 155, vi_lr_MoverWidth := 80);<br>
  FOR un_Module := 1 TO 6 DO<br>
      fb_Idh.m_SetModule(vi_un_Module := un_Module, vi_e_Kind := E_VisuModuleKind.STRAIGHT);<br>
  END_FOR<br>
  fb_Idh.m_SetFinger(vi_un_Finger := 1, vi_lr_Diameter := 40, vi_lr_Height := 50);<br>
  fb_Idh.m_SetZone(vi_un_Zone := 1, vi_udn_ConveyorId := 3, vi_lr_Start := 1100, vi_lr_End := 2600);<br>
  fb_Idh.m_SetZPosition(lr_ZAxisActual);<br>
  fb_Idh.m_SetMoverCount(4);<br>
  fb_Idh.m_SetMover(vi_un_Index := 0, vi_udn_Id := 1, vi_lr_Position := ..., vi_lr_X := ..., vi_FingerStates := Mover1Fingers);<br>
Only actual values are reported; tool rotations (e.g. C) show only through the finger poses, absolute in the MCS.<br>
The config methods may be called every cycle; the config version only changes when a value does.<br>
*****************************************************************************************************<br>
OUTPUT VALUES:<br>
vo_Visu is the contract structure the gateway reads at the path given to m_Register. Do not write it.<br>
*****************************************************************************************************<br>
VERSION         ¦ DATE       ¦ NAME      ¦ CHANGE<br>
Syn_Visu 3.0.0  ¦ 2026-10-31 ¦ J.Willner ¦ Naming and layout after the TCAT programming guideline<br>
Syn_Visu 4.0.0  ¦ 2026-11-01 ¦ J.Willner ¦ Zones and fingers from _FB_VisuRobot; m_SetZone by index, no kind<br>
Syn_Visu 5.0.0  ¦ 2026-11-01 ¦ J.Willner ¦ Track of modules from _FB_VisuXtsTrack (m_SetModule)<br>
****************************************************************************************************)
FUNCTION_BLOCK _FB_VisuXtsGantry EXTENDS _FB_VisuXtsTrack
VAR_OUTPUT
	vo_Visu								: ST_VisuXtsGantry;	// contract structure read by the gateway
END_VAR

(****************************************************************************************************<br>
© Syntegon Group.<br>
All rights reserved, also regarding any disposal, exploitation, reproduction, editing, distribution,<br>
as well as in the event of applications for industrial property rights.<br>
*****************************************************************************************************<br>
DESCRIPTION:<br>
Takes over vio_New and increments the config version if it differs from the current config. TRUE if changed.<br>
****************************************************************************************************)
METHOD PRIVATE m_ApplyConfig : BOOL
VAR_IN_OUT
	vio_New								: ST_VisuXtsGantryConfig;
END_VAR
m_ApplyConfig := Tc2_System.MEMCMP(ADR(vio_New), ADR(vo_Visu.stConfig), SIZEOF(vio_New)) <> 0;
IF m_ApplyConfig THEN
	vo_Visu.stConfig := vio_New;
	m_NotifyConfigChanged();
END_IF
END_METHOD

(****************************************************************************************************<br>
© Syntegon Group.<br>
All rights reserved, also regarding any disposal, exploitation, reproduction, editing, distribution,<br>
as well as in the event of applications for industrial property rights.<br>
*****************************************************************************************************<br>
DESCRIPTION:<br>
Manifest type: XTS gantry.<br>
****************************************************************************************************)
METHOD PROTECTED m_ComponentType : E_VisuComponentType
m_ComponentType := E_VisuComponentType.XTS_GANTRY;
END_METHOD

(****************************************************************************************************<br>
© Syntegon Group.<br>
All rights reserved, also regarding any disposal, exploitation, reproduction, editing, distribution,<br>
as well as in the event of applications for industrial property rights.<br>
*****************************************************************************************************<br>
DESCRIPTION:<br>
Sets pose, strokes, gripper offsets and mover size; the track comes from m_SetModule. TRUE if anything changed.<br>
****************************************************************************************************)
METHOD m_Configure : BOOL
VAR_INPUT
	vi_Pose								: ST_VisuPose;	// MCS, track start on top of the movers with Z = 0
	vi_lr_XMin							: LREAL;	// [mm]
	vi_lr_XMax							: LREAL;	// [mm]
	vi_lr_ZMin							: LREAL;	// [mm]
	vi_lr_ZMax							: LREAL;	// [mm]
	vi_lr_ToolOffsetX					: LREAL;	// [mm] gripper flange ahead of the X axis zero
	vi_lr_ToolOffsetZ					: LREAL;	// [mm] gripper flange relative to the mover top (below: negative)
	vi_lr_MoverLength					: LREAL;	// [mm] along the track
	vi_lr_MoverWidth					: LREAL;	// [mm]
END_VAR
VAR
	TempNew								: ST_VisuXtsGantryConfig;
END_VAR
TempNew := vo_Visu.stConfig;
TempNew.stPose := vi_Pose;
TempNew.fXMin := vi_lr_XMin;
TempNew.fXMax := vi_lr_XMax;
TempNew.fZMin := vi_lr_ZMin;
TempNew.fZMax := vi_lr_ZMax;
TempNew.fToolOffsetX := vi_lr_ToolOffsetX;
TempNew.fToolOffsetZ := vi_lr_ToolOffsetZ;
TempNew.fMoverLength := vi_lr_MoverLength;
TempNew.fMoverWidth := vi_lr_MoverWidth;
m_Configure := m_ApplyConfig(TempNew);
END_METHOD

(****************************************************************************************************<br>
© Syntegon Group.<br>
All rights reserved, also regarding any disposal, exploitation, reproduction, editing, distribution,<br>
as well as in the event of applications for industrial property rights.<br>
*****************************************************************************************************<br>
DESCRIPTION:<br>
The fingers of every mover's gripper for _FB_VisuRobot.m_SetFinger and m_ClearFingers.<br>
****************************************************************************************************)
METHOD PROTECTED m_Fingers : BOOL
VAR_OUTPUT
	vo_p_Count							: POINTER TO UINT;
	vo_p_Fingers						: POINTER TO ARRAY[0..VISU_GlobalConst_Param.VISU_un_MAX_FINGERS - 1] OF ST_VisuFinger;
END_VAR
vo_p_Count := ADR(vo_Visu.stConfig.nFingerCount);
vo_p_Fingers := ADR(vo_Visu.stConfig.aFingers);
m_Fingers := TRUE;
END_METHOD

(****************************************************************************************************<br>
© Syntegon Group.<br>
All rights reserved, also regarding any disposal, exploitation, reproduction, editing, distribution,<br>
as well as in the event of applications for industrial property rights.<br>
*****************************************************************************************************<br>
DESCRIPTION:<br>
The gantry's track modules for _FB_VisuXtsTrack.m_SetModule and m_ClearModules.<br>
****************************************************************************************************)
METHOD PROTECTED m_Modules : BOOL
VAR_OUTPUT
	vo_p_Count							: POINTER TO UINT;
	vo_p_Modules						: POINTER TO ARRAY[0..VISU_GlobalConst_Param.VISU_un_MAX_MODULES - 1] OF ST_VisuTrackModule;
	vo_p_States							: POINTER TO ARRAY[0..VISU_GlobalConst_Param.VISU_un_MAX_MODULES - 1] OF ST_VisuTrackModuleState;
END_VAR
vo_p_Count := ADR(vo_Visu.stConfig.nModuleCount);
vo_p_Modules := ADR(vo_Visu.stConfig.aModules);
vo_p_States := ADR(vo_Visu.stState.aModuleStates);
m_Modules := TRUE;
END_METHOD

(****************************************************************************************************<br>
© Syntegon Group.<br>
All rights reserved, also regarding any disposal, exploitation, reproduction, editing, distribution,<br>
as well as in the event of applications for industrial property rights.<br>
*****************************************************************************************************<br>
DESCRIPTION:<br>
Sets or clears the fault of the whole gantry: drawn red with the message while active. Faults of single<br>
movers go through m_SetMover. The fault stays until it is cleared with m_SetFault(vi_b_Active := FALSE,<br>
vi_str_Message := ''). TRUE.<br>
****************************************************************************************************)
METHOD m_SetFault : BOOL
VAR_INPUT
	vi_b_Active							: BOOL;	// TRUE: fault active
	vi_str_Message						: STRING(80);	// shown to the operator; empty shows 'Fault'
END_VAR
vo_Visu.stState.stFault.bActive := vi_b_Active;
vo_Visu.stState.stFault.sMessage := vi_str_Message;
m_SetFault := TRUE;
END_METHOD

(****************************************************************************************************<br>
© Syntegon Group.<br>
All rights reserved, also regarding any disposal, exploitation, reproduction, editing, distribution,<br>
as well as in the event of applications for industrial property rights.<br>
*****************************************************************************************************<br>
DESCRIPTION:<br>
Reports one mover (actual values) at entry vi_un_Index and marks it valid. Call once per cycle per mover.<br>
*****************************************************************************************************<br>
OUTPUT VALUES:<br>
FALSE if vi_un_Index is outside the mover count set by m_SetMoverCount.<br>
****************************************************************************************************)
METHOD m_SetMover : BOOL
VAR_INPUT
	vi_un_Index							: UINT;	// [-] 0..m_SetMoverCount - 1
	vi_udn_Id							: UDINT;	// [-] unique within the gantry, > 0
	vi_lr_Position						: LREAL;	// [mm] along the track
	vi_lr_X								: LREAL;	// [mm] X axis
	vi_b_GripperActive					: BOOL;	// used only when no fingers are configured
	(* Finger poses absolute in the MCS and grip states, index 0 = finger 1; entries beyond the finger count are ignored. *)
	vi_FingerStates						: ARRAY[0..VISU_GlobalConst_Param.VISU_un_MAX_FINGERS - 1] OF ST_VisuFingerState;
	vi_b_Fault							: BOOL := FALSE;	// TRUE: this mover is in a fault
	vi_str_FaultMessage					: STRING(80) := '';	// shown to the operator; empty shows 'Fault'
END_VAR
m_SetMover := vi_un_Index < vo_Visu.stState.nMoverCount;
IF m_SetMover THEN
	vo_Visu.stState.aMovers[vi_un_Index].nId := vi_udn_Id;
	vo_Visu.stState.aMovers[vi_un_Index].bValid := TRUE;
	vo_Visu.stState.aMovers[vi_un_Index].fPosition := vi_lr_Position;
	vo_Visu.stState.aMovers[vi_un_Index].fX := vi_lr_X;
	vo_Visu.stState.aMovers[vi_un_Index].bGripperActive := vi_b_GripperActive;
	vo_Visu.stState.aMovers[vi_un_Index].aFingerStates := vi_FingerStates;
	vo_Visu.stState.aMovers[vi_un_Index].stFault.bActive := vi_b_Fault;
	vo_Visu.stState.aMovers[vi_un_Index].stFault.sMessage := vi_str_FaultMessage;
	vo_Visu.stState.nTimestamp := m_DcTime();
END_IF
END_METHOD

(****************************************************************************************************<br>
© Syntegon Group.<br>
All rights reserved, also regarding any disposal, exploitation, reproduction, editing, distribution,<br>
as well as in the event of applications for industrial property rights.<br>
*****************************************************************************************************<br>
DESCRIPTION:<br>
Sets how many mover entries are evaluated (limited to VISU_GlobalConst_Param.VISU_un_MAX_MOVERS); entries<br>
beyond are invalidated. TRUE if vi_un_Count fitted.<br>
****************************************************************************************************)
METHOD m_SetMoverCount : BOOL
VAR_INPUT
	vi_un_Count							: UINT;	// [-] movers
END_VAR
VAR
	un_TempIndex						: UINT;
END_VAR
m_SetMoverCount := vi_un_Count <= VISU_GlobalConst_Param.VISU_un_MAX_MOVERS;
vo_Visu.stState.nMoverCount := MIN(vi_un_Count, VISU_GlobalConst_Param.VISU_un_MAX_MOVERS);
FOR un_TempIndex := vo_Visu.stState.nMoverCount TO VISU_GlobalConst_Param.VISU_un_MAX_MOVERS - 1 DO
	vo_Visu.stState.aMovers[un_TempIndex].bValid := FALSE;
END_FOR
END_METHOD

(****************************************************************************************************<br>
© Syntegon Group.<br>
All rights reserved, also regarding any disposal, exploitation, reproduction, editing, distribution,<br>
as well as in the event of applications for industrial property rights.<br>
*****************************************************************************************************<br>
DESCRIPTION:<br>
Moves the gantry's shown coordinate system (origin triad, local measuring coordinates) away from the track<br>
start (stPose), in the gantry's local frame. Geometry and mover positions stay relative to stPose.<br>
TRUE if anything changed.<br>
****************************************************************************************************)
METHOD m_SetOriginShift : BOOL
VAR_INPUT
	vi_lr_X								: LREAL;	// [mm] along the gantry's local X
	vi_lr_Y								: LREAL := 0;	// [mm] along the track (local Y)
	vi_lr_Z								: LREAL := 0;	// [mm] along the gantry's local Z
END_VAR
VAR
	TempNew								: ST_VisuXtsGantryConfig;
END_VAR
TempNew := vo_Visu.stConfig;
TempNew.stOriginShift.fX := vi_lr_X;
TempNew.stOriginShift.fY := vi_lr_Y;
TempNew.stOriginShift.fZ := vi_lr_Z;
m_SetOriginShift := m_ApplyConfig(TempNew);
END_METHOD

(****************************************************************************************************<br>
© Syntegon Group.<br>
All rights reserved, also regarding any disposal, exploitation, reproduction, editing, distribution,<br>
as well as in the event of applications for industrial property rights.<br>
*****************************************************************************************************<br>
DESCRIPTION:<br>
Reports the common Z axis (actual value). Call once per cycle; it also stamps the state with the cycle's DC time.<br>
****************************************************************************************************)
METHOD m_SetZPosition : BOOL
VAR_INPUT
	vi_lr_Z								: LREAL;	// [mm]
END_VAR
vo_Visu.stState.fZ := vi_lr_Z;
vo_Visu.stState.nTimestamp := m_DcTime();
m_SetZPosition := TRUE;
END_METHOD

(****************************************************************************************************<br>
© Syntegon Group.<br>
All rights reserved, also regarding any disposal, exploitation, reproduction, editing, distribution,<br>
as well as in the event of applications for industrial property rights.<br>
*****************************************************************************************************<br>
DESCRIPTION:<br>
The gantry's zones for _FB_VisuZoneComponent.m_SetZone and m_ClearZones.<br>
****************************************************************************************************)
METHOD PROTECTED m_Zones : BOOL
VAR_OUTPUT
	vo_p_Count							: POINTER TO UINT;
	vo_p_Zones							: POINTER TO ARRAY[0..VISU_GlobalConst_Param.VISU_un_MAX_ZONES - 1] OF ST_VisuZone;
END_VAR
vo_p_Count := ADR(vo_Visu.stConfig.nZoneCount);
vo_p_Zones := ADR(vo_Visu.stConfig.aZones);
m_Zones := TRUE;
END_METHOD

END_FUNCTION_BLOCK

// POUs/_FB_VisuXtsTrack
(****************************************************************************************************<br>
© Syntegon Group.<br>
All rights reserved, also regarding any disposal, exploitation, reproduction, editing, distribution,<br>
as well as in the event of applications for industrial property rights.<br>
*****************************************************************************************************<br>
DESCRIPTION:<br>
Base of the XTS kinematics (XTS gantry, XTS loop): a robot whose movers run along a track of XTS motor<br>
modules, m_SetModule, m_ClearModules, m_SetModuleFault and m_TrackLength. The track is a chain of modules in the order the movers<br>
run along it, each starting where the one before it ends: STRAIGHT, or a quarter curve CURVE_LEFT or CURVE_RIGHT.<br>
A derived FB tells where its modules lie through m_Modules. Not used directly.<br>
*****************************************************************************************************<br>
VERSION         ¦ DATE       ¦ NAME      ¦ CHANGE<br>
Syn_Visu 5.0.0  ¦ 2026-11-01 ¦ J.Willner ¦ New: XTS tracks of track modules, a fault per module<br>
****************************************************************************************************)
FUNCTION_BLOCK ABSTRACT _FB_VisuXtsTrack EXTENDS _FB_VisuRobot

(****************************************************************************************************<br>
© Syntegon Group.<br>
All rights reserved, also regarding any disposal, exploitation, reproduction, editing, distribution,<br>
as well as in the event of applications for industrial property rights.<br>
*****************************************************************************************************<br>
DESCRIPTION:<br>
Removes all track modules. TRUE if there were any.<br>
****************************************************************************************************)
METHOD m_ClearModules : BOOL
VAR
	p_TempCount							: POINTER TO UINT;
	p_TempModules						: POINTER TO ARRAY[0..VISU_GlobalConst_Param.VISU_un_MAX_MODULES - 1] OF ST_VisuTrackModule;
	TempEmpty							: ST_VisuTrackModule;
	un_TempIndex						: UINT;
END_VAR
m_ClearModules := FALSE;
m_Modules(vo_p_Count => p_TempCount, vo_p_Modules => p_TempModules);
IF p_TempCount = 0 OR p_TempModules = 0 THEN
	RETURN;
END_IF
m_ClearModules := p_TempCount^ > 0;
FOR un_TempIndex := 0 TO VISU_GlobalConst_Param.VISU_un_MAX_MODULES - 1 DO
	p_TempModules^[un_TempIndex] := TempEmpty;
END_FOR
p_TempCount^ := 0;
IF m_ClearModules THEN
	m_NotifyConfigChanged();
END_IF
END_METHOD

(****************************************************************************************************<br>
© Syntegon Group.<br>
All rights reserved, also regarding any disposal, exploitation, reproduction, editing, distribution,<br>
as well as in the event of applications for industrial property rights.<br>
*****************************************************************************************************<br>
DESCRIPTION:<br>
Where the track modules lie in the derived FB's contract structure: vo_p_Count points to its nModuleCount,<br>
vo_p_Modules to its aModules, vo_p_States to its state's aModuleStates.<br>
****************************************************************************************************)
METHOD PROTECTED ABSTRACT m_Modules : BOOL
VAR_OUTPUT
	vo_p_Count							: POINTER TO UINT;
	vo_p_Modules						: POINTER TO ARRAY[0..VISU_GlobalConst_Param.VISU_un_MAX_MODULES - 1] OF ST_VisuTrackModule;
	vo_p_States							: POINTER TO ARRAY[0..VISU_GlobalConst_Param.VISU_un_MAX_MODULES - 1] OF ST_VisuTrackModuleState;
END_VAR
END_METHOD

(****************************************************************************************************<br>
© Syntegon Group.<br>
All rights reserved, also regarding any disposal, exploitation, reproduction, editing, distribution,<br>
as well as in the event of applications for industrial property rights.<br>
*****************************************************************************************************<br>
DESCRIPTION:<br>
Sets track module vi_un_Module (1-based, in the order the movers run along the track): it starts where module<br>
vi_un_Module - 1 ends. The module count grows to vi_un_Module; set the modules in order. Track positions count<br>
from the start of module 1. The config version only changes when a value does.<br>
*****************************************************************************************************<br>
OUTPUT VALUES:<br>
FALSE for vi_un_Module outside 1..VISU_GlobalConst_Param.VISU_un_MAX_MODULES.<br>
****************************************************************************************************)
METHOD m_SetModule : BOOL
VAR_INPUT
	vi_un_Module						: UINT;	// [-] 1-based
	vi_e_Kind							: E_VisuModuleKind;	// straight, or a quarter curve to the left or right
	vi_lr_Length						: LREAL := VISU_GlobalConst.VISU_lr_XTS_MODULE_LENGTH;	// [mm] along the track
END_VAR
VAR
	p_TempCount							: POINTER TO UINT;
	p_TempModules						: POINTER TO ARRAY[0..VISU_GlobalConst_Param.VISU_un_MAX_MODULES - 1] OF ST_VisuTrackModule;
END_VAR
m_SetModule := FALSE;
IF vi_un_Module = 0 OR vi_un_Module > VISU_GlobalConst_Param.VISU_un_MAX_MODULES THEN
	RETURN;
END_IF
m_Modules(vo_p_Count => p_TempCount, vo_p_Modules => p_TempModules);
IF p_TempCount = 0 OR p_TempModules = 0 THEN
	RETURN;
END_IF
(* Compared member by member: the padding after eKind is not part of the value. *)
IF vi_un_Module > p_TempCount^
OR p_TempModules^[vi_un_Module - 1].eKind <> vi_e_Kind
OR p_TempModules^[vi_un_Module - 1].fLength <> vi_lr_Length
THEN
	p_TempModules^[vi_un_Module - 1].eKind := vi_e_Kind;
	p_TempModules^[vi_un_Module - 1].fLength := vi_lr_Length;
	p_TempCount^ := MAX(p_TempCount^, vi_un_Module);
	m_NotifyConfigChanged();
END_IF
m_SetModule := TRUE;
END_METHOD

(****************************************************************************************************<br>
© Syntegon Group.<br>
All rights reserved, also regarding any disposal, exploitation, reproduction, editing, distribution,<br>
as well as in the event of applications for industrial property rights.<br>
*****************************************************************************************************<br>
DESCRIPTION:<br>
Reports the fault of track module vi_un_Module (1-based, as in m_SetModule), e.g. an overtemperature of that<br>
motor module. The visualisation draws the module red with the message above it. Call it every cycle with the<br>
module's current state; vi_b_Fault = FALSE clears it.<br>
*****************************************************************************************************<br>
OUTPUT VALUES:<br>
FALSE for vi_un_Module outside 1..VISU_GlobalConst_Param.VISU_un_MAX_MODULES.<br>
****************************************************************************************************)
METHOD m_SetModuleFault : BOOL
VAR_INPUT
	vi_un_Module						: UINT;	// [-] 1-based
	vi_b_Fault							: BOOL;	// TRUE: this module is in a fault
	vi_str_FaultMessage					: STRING(80) := '';	// shown to the operator; empty shows 'Fault'
END_VAR
VAR
	p_TempCount							: POINTER TO UINT;
	p_TempModules						: POINTER TO ARRAY[0..VISU_GlobalConst_Param.VISU_un_MAX_MODULES - 1] OF ST_VisuTrackModule;
	p_TempStates						: POINTER TO ARRAY[0..VISU_GlobalConst_Param.VISU_un_MAX_MODULES - 1] OF ST_VisuTrackModuleState;
END_VAR
m_SetModuleFault := FALSE;
IF vi_un_Module = 0 OR vi_un_Module > VISU_GlobalConst_Param.VISU_un_MAX_MODULES THEN
	RETURN;
END_IF
m_Modules(vo_p_Count => p_TempCount, vo_p_Modules => p_TempModules, vo_p_States => p_TempStates);
IF p_TempStates = 0 THEN
	RETURN;
END_IF
p_TempStates^[vi_un_Module - 1].stFault.bActive := vi_b_Fault;
p_TempStates^[vi_un_Module - 1].stFault.sMessage := vi_str_FaultMessage;
m_SetModuleFault := TRUE;
END_METHOD

(****************************************************************************************************<br>
© Syntegon Group.<br>
All rights reserved, also regarding any disposal, exploitation, reproduction, editing, distribution,<br>
as well as in the event of applications for industrial property rights.<br>
*****************************************************************************************************<br>
DESCRIPTION:<br>
Length of the track along its modules, [mm]: the range of track positions (on an XTS loop the perimeter).<br>
****************************************************************************************************)
METHOD m_TrackLength : LREAL
VAR
	p_TempCount							: POINTER TO UINT;
	p_TempModules						: POINTER TO ARRAY[0..VISU_GlobalConst_Param.VISU_un_MAX_MODULES - 1] OF ST_VisuTrackModule;
	un_TempIndex						: UINT;
END_VAR
m_TrackLength := 0;
m_Modules(vo_p_Count => p_TempCount, vo_p_Modules => p_TempModules);
IF p_TempCount = 0 OR p_TempModules = 0 THEN
	RETURN;
END_IF
FOR un_TempIndex := 1 TO MIN(p_TempCount^, VISU_GlobalConst_Param.VISU_un_MAX_MODULES) DO
	m_TrackLength := m_TrackLength + p_TempModules^[un_TempIndex - 1].fLength;
END_FOR
END_METHOD

END_FUNCTION_BLOCK

// POUs/_FB_VisuXtsLoop
(****************************************************************************************************<br>
© Syntegon Group.<br>
All rights reserved, also regarding any disposal, exploitation, reproduction, editing, distribution,<br>
as well as in the event of applications for industrial property rights.<br>
*****************************************************************************************************<br>
DESCRIPTION:<br>
One visualised XTS loop (e.g. Fxx): movers circulating on a closed track of XTS motor modules, e.g. two<br>
straights joined at each end by two CURVE_LEFT modules, standing in the local X-Z plane.<br>
Typical cycle:<br>
  fb_Fxx.m_Register(vio_Manifest := GVL_Visu.stManifest, vi_udn_Id := 20, vi_str_Name := 'Fxx',<br>
      vi_str_Path := 'MAIN.fb_Fxx.vo_Visu');<br>
  fb_Fxx.m_Configure(vi_Pose := LoopPose, vi_lr_ToolOffset := 120, vi_lr_MoverLength := 100,<br>
      vi_lr_MoverWidth := 60);<br>
  fb_Fxx.m_SetModule(vi_un_Module := 1, vi_e_Kind := E_VisuModuleKind.STRAIGHT); and so on, in order<br>
  fb_Fxx.m_SetFinger(vi_un_Finger := 1, vi_lr_Diameter := 40, vi_lr_Height := 50);<br>
  fb_Fxx.m_SetZone(vi_un_Zone := 1, vi_udn_ConveyorId := 2, vi_lr_Start := 2200, vi_lr_End := 2800);<br>
  fb_Fxx.m_SetMoverCount(12);<br>
  fb_Fxx.m_SetMover(vi_un_Index := 0, vi_udn_Id := 1, vi_lr_Position := ..., vi_FingerStates := Mover1Fingers);<br>
Positions run along the loop from the start of module 1 in the conveying direction (0..m_TrackLength()).<br>
The config methods may be called every cycle; the config version only changes when a value does.<br>
*****************************************************************************************************<br>
OUTPUT VALUES:<br>
vo_Visu is the contract structure the gateway reads at the path given to m_Register. Do not write it.<br>
*****************************************************************************************************<br>
VERSION         ¦ DATE       ¦ NAME      ¦ CHANGE<br>
Syn_Visu 3.0.0  ¦ 2026-10-31 ¦ J.Willner ¦ Naming and layout after the TCAT programming guideline<br>
Syn_Visu 4.0.0  ¦ 2026-11-01 ¦ J.Willner ¦ Zones and fingers from _FB_VisuRobot; m_SetZone by index, no kind<br>
Syn_Visu 5.0.0  ¦ 2026-11-01 ¦ J.Willner ¦ Track of modules from _FB_VisuXtsTrack; m_Perimeter is m_TrackLength<br>
****************************************************************************************************)
FUNCTION_BLOCK _FB_VisuXtsLoop EXTENDS _FB_VisuXtsTrack
VAR_OUTPUT
	vo_Visu								: ST_VisuXtsLoop;	// contract structure read by the gateway
END_VAR

(****************************************************************************************************<br>
© Syntegon Group.<br>
All rights reserved, also regarding any disposal, exploitation, reproduction, editing, distribution,<br>
as well as in the event of applications for industrial property rights.<br>
*****************************************************************************************************<br>
DESCRIPTION:<br>
Takes over vio_New and increments the config version if it differs from the current config. TRUE if changed.<br>
****************************************************************************************************)
METHOD PRIVATE m_ApplyConfig : BOOL
VAR_IN_OUT
	vio_New								: ST_VisuXtsLoopConfig;
END_VAR
m_ApplyConfig := Tc2_System.MEMCMP(ADR(vio_New), ADR(vo_Visu.stConfig), SIZEOF(vio_New)) <> 0;
IF m_ApplyConfig THEN
	vo_Visu.stConfig := vio_New;
	m_NotifyConfigChanged();
END_IF
END_METHOD

(****************************************************************************************************<br>
© Syntegon Group.<br>
All rights reserved, also regarding any disposal, exploitation, reproduction, editing, distribution,<br>
as well as in the event of applications for industrial property rights.<br>
*****************************************************************************************************<br>
DESCRIPTION:<br>
Manifest type: XTS loop.<br>
****************************************************************************************************)
METHOD PROTECTED m_ComponentType : E_VisuComponentType
m_ComponentType := E_VisuComponentType.XTS_LOOP;
END_METHOD

(****************************************************************************************************<br>
© Syntegon Group.<br>
All rights reserved, also regarding any disposal, exploitation, reproduction, editing, distribution,<br>
as well as in the event of applications for industrial property rights.<br>
*****************************************************************************************************<br>
DESCRIPTION:<br>
Sets pose, tool offset and mover size; the track comes from m_SetModule. TRUE if anything changed.<br>
****************************************************************************************************)
METHOD m_Configure : BOOL
VAR_INPUT
	vi_Pose								: ST_VisuPose;	// MCS, start of module 1; the loop stands in the local X-Z plane
	vi_lr_ToolOffset					: LREAL;	// [mm] tool point outwards from the track
	vi_lr_MoverLength					: LREAL;	// [mm] along the track
	vi_lr_MoverWidth					: LREAL;	// [mm]
END_VAR
VAR
	TempNew								: ST_VisuXtsLoopConfig;
END_VAR
TempNew := vo_Visu.stConfig;
TempNew.stPose := vi_Pose;
TempNew.fToolOffset := vi_lr_ToolOffset;
TempNew.fMoverLength := vi_lr_MoverLength;
TempNew.fMoverWidth := vi_lr_MoverWidth;
m_Configure := m_ApplyConfig(TempNew);
END_METHOD

(****************************************************************************************************<br>
© Syntegon Group.<br>
All rights reserved, also regarding any disposal, exploitation, reproduction, editing, distribution,<br>
as well as in the event of applications for industrial property rights.<br>
*****************************************************************************************************<br>
DESCRIPTION:<br>
The fingers of every mover's gripper for _FB_VisuRobot.m_SetFinger and m_ClearFingers.<br>
****************************************************************************************************)
METHOD PROTECTED m_Fingers : BOOL
VAR_OUTPUT
	vo_p_Count							: POINTER TO UINT;
	vo_p_Fingers						: POINTER TO ARRAY[0..VISU_GlobalConst_Param.VISU_un_MAX_FINGERS - 1] OF ST_VisuFinger;
END_VAR
vo_p_Count := ADR(vo_Visu.stConfig.nFingerCount);
vo_p_Fingers := ADR(vo_Visu.stConfig.aFingers);
m_Fingers := TRUE;
END_METHOD

(****************************************************************************************************<br>
© Syntegon Group.<br>
All rights reserved, also regarding any disposal, exploitation, reproduction, editing, distribution,<br>
as well as in the event of applications for industrial property rights.<br>
*****************************************************************************************************<br>
DESCRIPTION:<br>
The loop's track modules for _FB_VisuXtsTrack.m_SetModule and m_ClearModules.<br>
****************************************************************************************************)
METHOD PROTECTED m_Modules : BOOL
VAR_OUTPUT
	vo_p_Count							: POINTER TO UINT;
	vo_p_Modules						: POINTER TO ARRAY[0..VISU_GlobalConst_Param.VISU_un_MAX_MODULES - 1] OF ST_VisuTrackModule;
	vo_p_States							: POINTER TO ARRAY[0..VISU_GlobalConst_Param.VISU_un_MAX_MODULES - 1] OF ST_VisuTrackModuleState;
END_VAR
vo_p_Count := ADR(vo_Visu.stConfig.nModuleCount);
vo_p_Modules := ADR(vo_Visu.stConfig.aModules);
vo_p_States := ADR(vo_Visu.stState.aModuleStates);
m_Modules := TRUE;
END_METHOD

(****************************************************************************************************<br>
© Syntegon Group.<br>
All rights reserved, also regarding any disposal, exploitation, reproduction, editing, distribution,<br>
as well as in the event of applications for industrial property rights.<br>
*****************************************************************************************************<br>
DESCRIPTION:<br>
Sets or clears the fault of the whole loop: drawn red with the message while active. Faults of single<br>
movers go through m_SetMover. The fault stays until it is cleared with m_SetFault(vi_b_Active := FALSE,<br>
vi_str_Message := ''). TRUE.<br>
****************************************************************************************************)
METHOD m_SetFault : BOOL
VAR_INPUT
	vi_b_Active							: BOOL;	// TRUE: fault active
	vi_str_Message						: STRING(80);	// shown to the operator; empty shows 'Fault'
END_VAR
vo_Visu.stState.stFault.bActive := vi_b_Active;
vo_Visu.stState.stFault.sMessage := vi_str_Message;
m_SetFault := TRUE;
END_METHOD

(****************************************************************************************************<br>
© Syntegon Group.<br>
All rights reserved, also regarding any disposal, exploitation, reproduction, editing, distribution,<br>
as well as in the event of applications for industrial property rights.<br>
*****************************************************************************************************<br>
DESCRIPTION:<br>
Reports one mover at entry vi_un_Index and marks it valid. Call once per cycle per mover.<br>
*****************************************************************************************************<br>
OUTPUT VALUES:<br>
FALSE if vi_un_Index is outside the mover count set by m_SetMoverCount.<br>
****************************************************************************************************)
METHOD m_SetMover : BOOL
VAR_INPUT
	vi_un_Index							: UINT;	// [-] 0..m_SetMoverCount - 1
	vi_udn_Id							: UDINT;	// [-] unique within the loop, > 0
	vi_lr_Position						: LREAL;	// [mm] along the loop from the start of module 1 (0..m_TrackLength())
	(* Finger poses absolute in the MCS and grip states, index 0 = finger 1; entries beyond the finger count are ignored. *)
	vi_FingerStates						: ARRAY[0..VISU_GlobalConst_Param.VISU_un_MAX_FINGERS - 1] OF ST_VisuFingerState;
	vi_b_Fault							: BOOL := FALSE;	// TRUE: this mover is in a fault
	vi_str_FaultMessage					: STRING(80) := '';	// shown to the operator; empty shows 'Fault'
END_VAR
m_SetMover := vi_un_Index < vo_Visu.stState.nMoverCount;
IF m_SetMover THEN
	vo_Visu.stState.aMovers[vi_un_Index].nId := vi_udn_Id;
	vo_Visu.stState.aMovers[vi_un_Index].bValid := TRUE;
	vo_Visu.stState.aMovers[vi_un_Index].fPosition := vi_lr_Position;
	vo_Visu.stState.aMovers[vi_un_Index].aFingerStates := vi_FingerStates;
	vo_Visu.stState.aMovers[vi_un_Index].stFault.bActive := vi_b_Fault;
	vo_Visu.stState.aMovers[vi_un_Index].stFault.sMessage := vi_str_FaultMessage;
	vo_Visu.stState.nTimestamp := m_DcTime();
END_IF
END_METHOD

(****************************************************************************************************<br>
© Syntegon Group.<br>
All rights reserved, also regarding any disposal, exploitation, reproduction, editing, distribution,<br>
as well as in the event of applications for industrial property rights.<br>
*****************************************************************************************************<br>
DESCRIPTION:<br>
Sets how many mover entries are evaluated (limited to VISU_GlobalConst_Param.VISU_un_MAX_MOVERS); entries<br>
beyond are invalidated. TRUE if vi_un_Count fitted.<br>
****************************************************************************************************)
METHOD m_SetMoverCount : BOOL
VAR_INPUT
	vi_un_Count							: UINT;	// [-] movers
END_VAR
VAR
	un_TempIndex						: UINT;
END_VAR
m_SetMoverCount := vi_un_Count <= VISU_GlobalConst_Param.VISU_un_MAX_MOVERS;
vo_Visu.stState.nMoverCount := MIN(vi_un_Count, VISU_GlobalConst_Param.VISU_un_MAX_MOVERS);
FOR un_TempIndex := vo_Visu.stState.nMoverCount TO VISU_GlobalConst_Param.VISU_un_MAX_MOVERS - 1 DO
	vo_Visu.stState.aMovers[un_TempIndex].bValid := FALSE;
END_FOR
END_METHOD

(****************************************************************************************************<br>
© Syntegon Group.<br>
All rights reserved, also regarding any disposal, exploitation, reproduction, editing, distribution,<br>
as well as in the event of applications for industrial property rights.<br>
*****************************************************************************************************<br>
DESCRIPTION:<br>
Moves the loop's shown coordinate system (origin triad, local measuring coordinates) away from the start of<br>
the lower straight (stPose), in the loop's local frame. Geometry and mover positions stay relative to stPose.<br>
TRUE if anything changed.<br>
****************************************************************************************************)
METHOD m_SetOriginShift : BOOL
VAR_INPUT
	vi_lr_X								: LREAL;	// [mm] along the lower straight (local X)
	vi_lr_Y								: LREAL := 0;	// [mm] along the loop's local Y
	vi_lr_Z								: LREAL := 0;	// [mm] along the loop's local Z
END_VAR
VAR
	TempNew								: ST_VisuXtsLoopConfig;
END_VAR
TempNew := vo_Visu.stConfig;
TempNew.stOriginShift.fX := vi_lr_X;
TempNew.stOriginShift.fY := vi_lr_Y;
TempNew.stOriginShift.fZ := vi_lr_Z;
m_SetOriginShift := m_ApplyConfig(TempNew);
END_METHOD

(****************************************************************************************************<br>
© Syntegon Group.<br>
All rights reserved, also regarding any disposal, exploitation, reproduction, editing, distribution,<br>
as well as in the event of applications for industrial property rights.<br>
*****************************************************************************************************<br>
DESCRIPTION:<br>
The loop's zones for _FB_VisuZoneComponent.m_SetZone and m_ClearZones.<br>
****************************************************************************************************)
METHOD PROTECTED m_Zones : BOOL
VAR_OUTPUT
	vo_p_Count							: POINTER TO UINT;
	vo_p_Zones							: POINTER TO ARRAY[0..VISU_GlobalConst_Param.VISU_un_MAX_ZONES - 1] OF ST_VisuZone;
END_VAR
vo_p_Count := ADR(vo_Visu.stConfig.nZoneCount);
vo_p_Zones := ADR(vo_Visu.stConfig.aZones);
m_Zones := TRUE;
END_METHOD

END_FUNCTION_BLOCK

// POUs/_FC_GetVersionSynVisu
(****************************************************************************************************<br>
© Syntegon Group.<br>
All rights reserved, also regarding any disposal, exploitation, reproduction, editing, distribution,<br>
as well as in the event of applications for industrial property rights.<br>
*****************************************************************************************************<br>
DESCRIPTION:<br>
Runtime-readable version of the Syn_Visu library.<br>
*****************************************************************************************************<br>
VERSION         ¦ DATE       ¦ NAME      ¦ CHANGE<br>
Syn_Visu 3.0.0  ¦ 2026-10-31 ¦ J.Willner ¦ Naming and layout after the TCAT programming guideline<br>
Syn_Visu 3.1.0  ¦ 2026-10-31 ¦ J.Willner ¦ Faults of components and XTS movers (protocol 8)<br>
Syn_Visu 3.2.0  ¦ 2026-10-31 ¦ J.Willner ¦ _FB_VisuConveyor.m_MoveProduct<br>
Syn_Visu 3.3.0  ¦ 2026-10-31 ¦ J.Willner ¦ Zone CCS offset, origin shift per component (protocol 9)<br>
Syn_Visu 3.4.0  ¦ 2026-11-01 ¦ J.Willner ¦ m_LatchProduct: product state and robot (PLACED onto outfeeds)<br>
Syn_Visu 3.5.0  ¦ 2026-11-01 ¦ J.Willner ¦ Product shapes: box, cylinder, rounded box (protocol 10)<br>
Syn_Visu 4.0.0  ¦ 2026-11-01 ¦ J.Willner ¦ Vision system, product sensor, zones without kind (protocol 11)<br>
Syn_Visu 5.0.0  ¦ 2026-11-01 ¦ J.Willner ¦ XTS tracks of track modules, a fault per module (protocol 12)<br>
Syn_Visu 5.1.0  ¦ 2026-11-01 ¦ J.Willner ¦ Manifest sLibraryVersion: the visualisation shows the library version<br>
Syn_Visu 6.0.0  ¦ 2026-11-01 ¦ J.Willner ¦ Generic product client (nLastClientId, ePreviousState), station (protocol 13)<br>
****************************************************************************************************)
FUNCTION _FC_GetVersionSynVisu : UINT
VAR_INPUT
	vi_n_VersionElement					: INT;	// [-] 1 = major, 2 = minor, 3 = revision
END_VAR

CASE vi_n_VersionElement OF
	1: _FC_GetVersionSynVisu := 6;
	2: _FC_GetVersionSynVisu := 0;
	3: _FC_GetVersionSynVisu := 0;
ELSE
	_FC_GetVersionSynVisu := 16#FFFF;
END_CASE

END_FUNCTION
